Universal Robots PolyScope program: universal_robots_robot_motion_script.urp

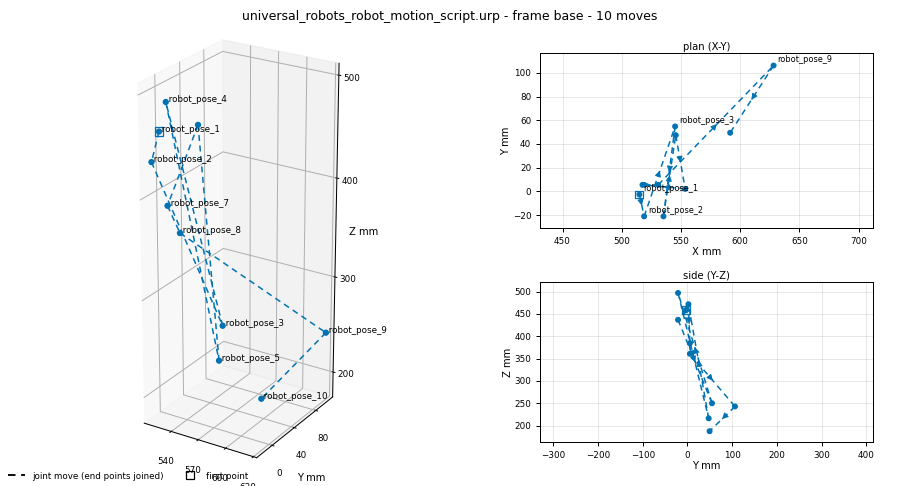
[picture p0: tool path of universal_robots_robot_motion_script.urp in frame base, 10 of 10 moves have a stored position in this frame; points joined in program order, loops and branches not executed]
Program universal_robots_robot_motion_script (installation=default directory=/programs/usbdisk createdIn=5.5.1 lastSavedIn=5.13.0 robotSerialNumber=20235500398)
Calibrated DH parameters: a=[0.000123, -0.269911, -0.358672, 0.000007, 0.000086, 0]; d=[0.162481, 303.203719, -198.264652, -104.805533, 0.099782, 0.099767]; alpha=[1.570424, -0.001084, -0.001515, 1.570177, -1.570736, 0]; deltaTheta=[0, -0.883345, 6.749397, 0.41713, 0, 0]
InitVariablesNode variables(variable(name=Counter, expression=0))
Robot Program (runOnlyOnce=false)
  'set image_counter to 0'
  Script: write_output_integer_register(24,0)
  'set start_capture to False'
  Script: write_output_boolean_register(64,False)
  SuppressedNode
    Wait DigitalInput pin=GP_bool_in[65]; digitalValue=1
  Wait Condition expression=read_input_boolean_register(65)
  Script: read_input_boolean_register(65)
  'Add, alter, or remove waypoints to calibrate'
  MoveJ speed 15 deg/s, acceleration 15 deg/s^2 (useActiveTCP=true) feature=Base
    Waypoint robot_pose_1: TCP in base x=514.911 y=-2.606 z=458.971 mm, rx=-0.6764 ry=2.9145 rz=-0.1502 rad; joints [15.975, -88.877, -97.62, -75.413, -276.232, 79.357] deg
    Call capture_hand_eye
    Waypoint robot_pose_2: TCP in base x=518.875 y=-21.086 z=436.72 mm, rx=-1.0277 ry=2.8103 rz=0.0126 rad; joints [12.252, -90.351, -99.453, -71.792, -268.461, 62.14] deg
    Call capture_hand_eye
    Waypoint robot_pose_3: TCP in base x=545.046 y=54.826 z=250.04 mm, rx=1.2149 ry=-2.7761 rz=0.3224 rad; joints [22.158, -104.762, -108.91, -61.489, -282.341, 65.367] deg
    Call capture_hand_eye
    Waypoint robot_pose_4: TCP in base x=535.184 y=-21.087 z=496.794 mm, rx=0.9249 ry=-2.7352 rz=0.2638 rad; joints [14.355, -96.376, -79.247, -107.628, -281.418, 68.302] deg
    Call capture_hand_eye
    Waypoint robot_pose_5: TCP in base x=545.586 y=47.414 z=216.419 mm, rx=0.7908 ry=-3.0119 rz=0.3288 rad; joints [21.323, -107.431, -112.289, -52.268, -281.982, 82.021] deg
    Call capture_hand_eye
    Waypoint robot_pose_6: TCP in base x=553.523 y=2.139 z=471.58 mm, rx=0.8586 ry=-2.9397 rz=0.0707 rad; joints [14.7, -96.987, -83.861, -93.565, -272.872, 72.215] deg
    Call capture_hand_eye
    Waypoint robot_pose_7: TCP in base x=517.49 y=5.485 z=384.653 mm, rx=-0.9337 ry=2.8471 rz=0.1368 rad; joints [14.428, -92.144, -105.34, -64.708, -264.369, 68.437] deg
    Call capture_hand_eye
    Waypoint robot_pose_8: TCP in base x=530.751 y=5.483 z=360.641 mm, rx=0.5138 ry=-2.8954 rz=0.185 rad; joints [16.307, -97.556, -98.049, -86.339, -275.976, 86.76] deg
    Call capture_hand_eye
    Waypoint robot_pose_9: TCP in base x=628.14 y=106.213 z=242.95 mm, rx=0.0642 ry=-2.915 rz=0.1564 rad; joints [21.909, -117.816, -88.599, -77.639, -271.335, 109.472] deg
    Call capture_hand_eye
    Waypoint robot_pose_10: TCP in base x=591.501 y=49.464 z=187.574 mm, rx=0.5846 ry=-3.0058 rz=0.0522 rad; joints [18.035, -115.708, -103.945, -55.079, -271.467, 85.987] deg
    Call capture_hand_eye
  'Calibration complete'
  SuppressedNode
    Set ExpressionOutput pin=GP_int_out[24]; expression=-1
  Script: write_output_integer_register(24,-1)
  Halt
SubProgram -> capture_hand_eye
SubProgram capture_hand_eye (keepSynchronizedWithDisk=false)
  Wait Sleep waitTime=2
  Counter := Counter+1
  SuppressedNode
    Set ExpressionOutput pin=GP_int_out[24]; expression=Counter
  Script: write_output_integer_register(24,Counter)
  SuppressedNode
    Set DigitalOutput pin=GP_bool_out[64]; digitalValue=1
  Script: write_output_boolean_register(64, True)
  Wait Condition expression=read_input_boolean_register(64)
  SuppressedNode
    Set DigitalOutput pin=GP_bool_out[64]; digitalValue=0
  Script: write_output_boolean_register(64, False)
